// TIA Portal V21 export
TagTable "T_V2"
  X_V2 :   (PLC tag "HMI_IF".SwOn, HMI_Connection_1, 100 ms)
